FUNCTION_BLOCK FB_PendantPreInitState EXTENDS FB_PendantState
VAR_INPUT
END_VAR
VAR_OUTPUT
END_VAR
VAR
END_VAR

METHOD FoundError : BOOL
pPendant^.SetState(pPendant^.fbPendantErrorState);
END_METHOD

METHOD InitCommand : BOOL
pPendant^.SetState(pPendant^.fbPendantInitState);
END_METHOD

PROPERTY StateID : STRING
GET
StateID := 'Pre Init State';
END_GET
END_PROPERTY

END_FUNCTION_BLOCK

(* stored: Version 1.1.0.1, ProductVersion 3.1.4024.15
   POU FB_PendantPreInitState: Id {79cdc163-ce8d-4317-a0b7-e539911b12eb}, SpecialFunc None
   Method FoundError: Id {068bbf7a-f119-4b44-9bb0-3b3f032c4a80}
   Method InitCommand: Id {0e339302-0e5c-4517-896c-4d890de71cf3}
   Property StateID: Id {bac1925c-c344-4e99-a865-978a2d14402e}
   Get Get: Id {fb8a5ea7-6134-4bcc-9c7e-949fd01d9f60} *)
